Fanuc KAREL source: KA00125.KL

PROGRAM KA00125
%NOLOCKGROUP
VAR
  SRC: ARRAY[2] OF BYTE
  DST: POSITION
BEGIN
  SRC[1] = 2
  DST = SRC[1]
END KA00125
